// SIMATIC S7-200 project (STEP 7-Micro/WIN), CPU 224XP CN REL 02.01

ORGANIZATION_BLOCK MAIN:OB1
TITLE=REALIZADO POR: BISMARK CHOQUE CHOQUE - REALIMENTACION DE ESTADOS
BEGIN
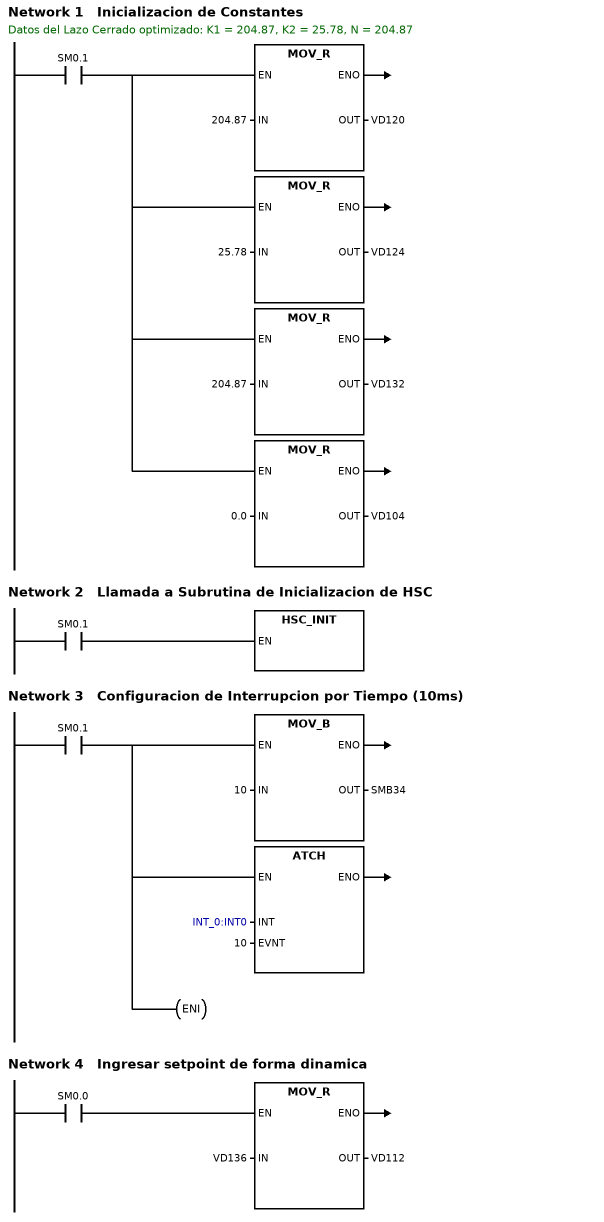
Network 1 //  Inicializacion de Constantes 
//  Datos del Lazo Cerrado optimizado: K1 = 204.87, K2 = 25.78, N = 204.87
// TU GANANCIA K1 (Posición)
// TU GANANCIA K2 (Velocidad)
// TU GANANCIA N (Pre-compensación calculada)
// Inicializar Pos_Anterior en 0.0
LD     SM0.1
MOVR   204.87, VD120
MOVR   25.78, VD124
MOVR   204.87, VD132
MOVR   0.0, VD104
Network 2 //  Llamada a Subrutina de Inicializacion de HSC
// Llamada a HSC_INIT
LD     SM0.1
CALL   HSC_INIT:SBR1
Network 3 //  Configuracion de Interrupcion por Tiempo (10ms)
// Intervalo de tiempo = 10 ms
// Asociar INT0 al evento de tiempo de SMB34
// Habilitar interrupciones globales
LD     SM0.1
MOVB   10, SMB34
ATCH   INT_0:INT0, 10
ENI
Network 4 //  Ingresar setpoint de forma dinamica
// Mover Setpoint desde VD136 a VD112
LD     SM0.0
MOVR   VD136, VD112
END_ORGANIZATION_BLOCK

SUBROUTINE_BLOCK HSC_INIT:SBR1
TITLE=
BEGIN
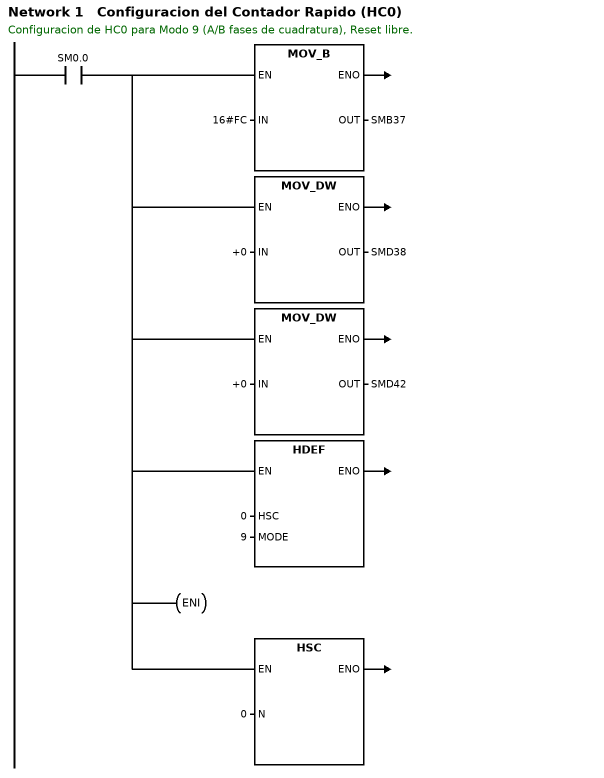
Network 1 //  Configuracion del Contador Rapido (HC0)
//  Configuracion de HC0 para Modo 9 (A/B fases de cuadratura), Reset libre.
// Control bits: Dirección arriba; escala 1X; habilitado
// Cargar valor actual en 0
// Cargar valor de preselección en 0
// Definir HC0 en Modo 9
// Asegurar habilitación de interrupciones
// Arrancar el contador rápido HC0
LD     SM0.0
MOVB   16#FC, SMB37
MOVD   +0, SMD38
MOVD   +0, SMD42
HDEF   0, 9
ENI
HSC    0
END_SUBROUTINE_BLOCK

INTERRUPT_BLOCK INT_0:INT0
TITLE=
BEGIN
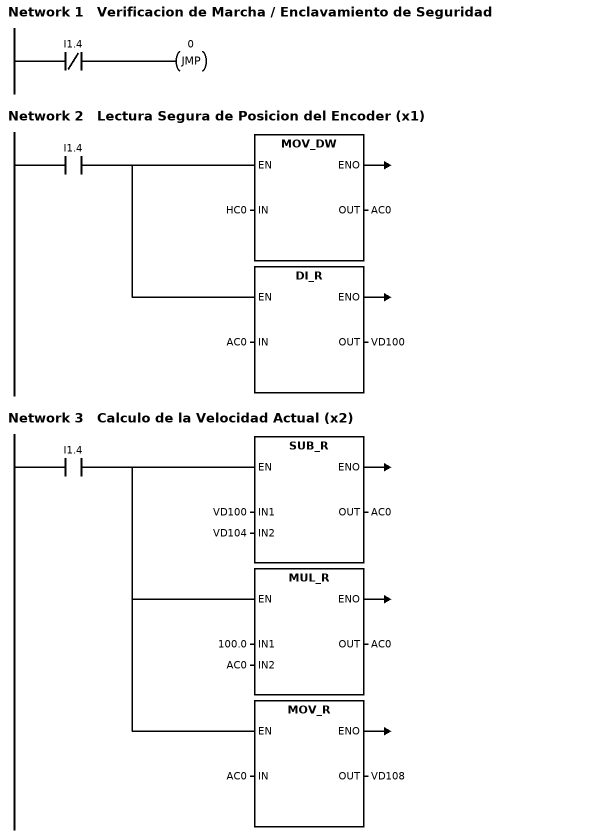
Network 1 //  Verificacion de Marcha / Enclavamiento de Seguridad
// Si I1.4 está desactivado (Emergencia/Stop)
// Salta directo a la parada segura (LBL 0)
LDN    I1.4
JMP    0
Network 2 //  Lectura Segura de Posicion del Encoder (x1)
// Leer cuentas acumuladas del hardware a AC0
// Convertir cuentas DINT a flotante REAL (x1)
LD     I1.4
MOVD   HC0, AC0
DTR    AC0, VD100
Network 3 //  Calculo de la Velocidad Actual (x2)
// Cuentas actuales
// Delta Posición = Cuentas_Actuales - Cuentas_Anteriores
// Delta_Pos / 0.01s equivale a multiplicar por 100.0
// Guardar en VD108 = Velocidad actual (x2)
LD     I1.4
MOVR   VD100, AC0
-R     VD104, AC0
*R     100.0, AC0
MOVR   AC0, VD108
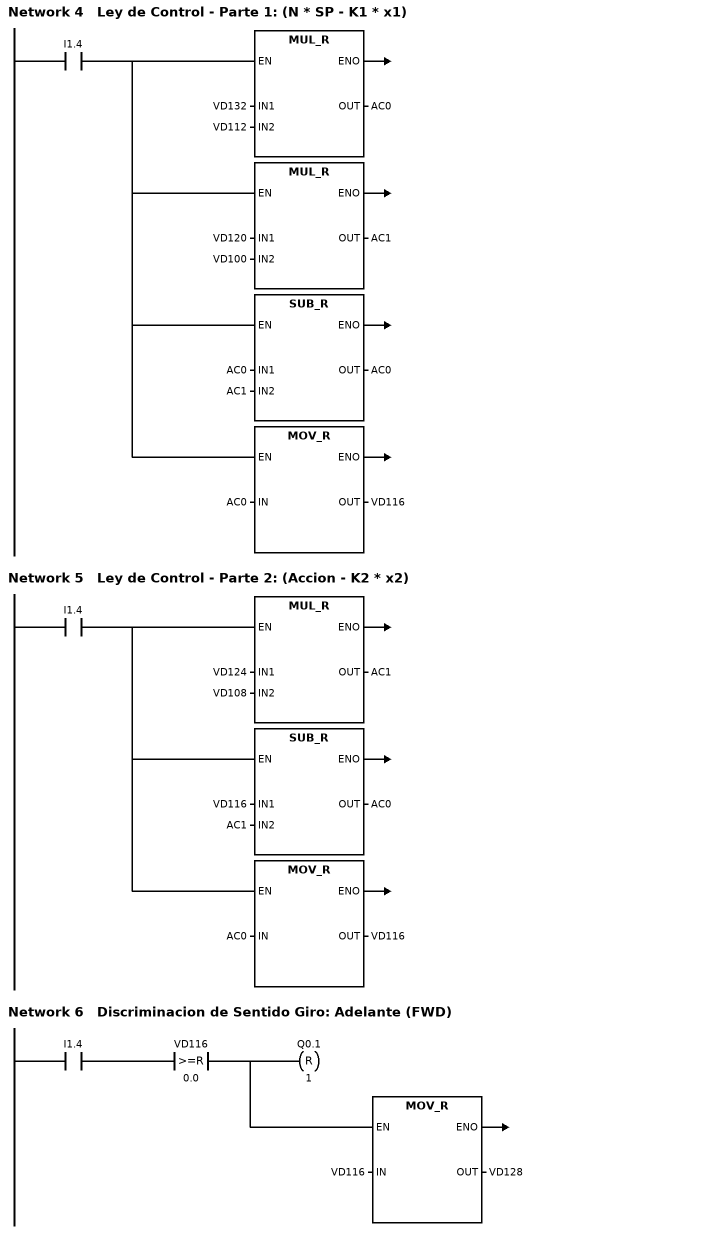
Network 4 //  Ley de Control - Parte 1: (N * SP - K1 * x1)
// Cargar N (204.87)
// AC0 = N * Setpoint
// Cargar K1 (204.87)
// AC1 = K1 * x1 (Posición)
// AC0 = (N * SP) - (K1 * x1)
// Almacenamiento intermedio
LD     I1.4
MOVR   VD132, AC0
*R     VD112, AC0
MOVR   VD120, AC1
*R     VD100, AC1
-R     AC1, AC0
MOVR   AC0, VD116
Network 5 //  Ley de Control - Parte 2: (Accion - K2 * x2)
// Cargar K2 (25.78)
// AC1 = K2 * x2 (Velocidad)
// Recuperar parte 1
// AC0 = (N * SP) - (K1 * x1) - (K2 * x2)
// VD116 = Acción de Control Final calculada (u)
LD     I1.4
MOVR   VD124, AC1
*R     VD108, AC1
MOVR   VD116, AC0
-R     AC1, AC0
MOVR   AC0, VD116
Network 6 //  Discriminacion de Sentido Giro: Adelante (FWD)
// Si u[k] es positiva o cero
// Desactivar salida de dirección reversa (Giro FWD)
// Guardar valor para magnitud |u|
LD     I1.4
AR>=   VD116, 0.0
R      Q0.1, 1
MOVR   VD116, VD128
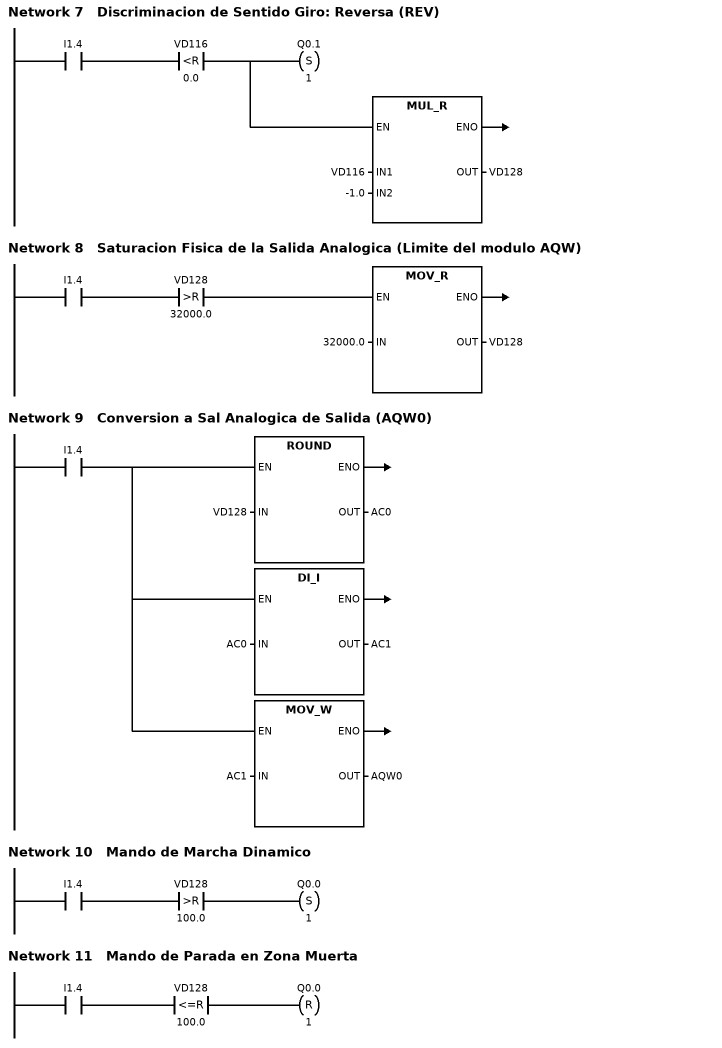
Network 7 //  Discriminacion de Sentido Giro: Reversa (REV)
// Si u[k] es negativa
// Activar salida física Q0.1 (Giro REV)
// Cargar u[k]
// Invertir signo para obtener valor absoluto |u|
LD     I1.4
AR<    VD116, 0.0
S      Q0.1, 1
MOVR   VD116, VD128
*R     -1.0, VD128
Network 8 //  Saturacion Fisica de la Salida Analogica (Limite del modulo AQW)
// Si excede el límite del módulo analógico de Siemens
// Recortar la acción a un máximo de 32000 unidades
LD     I1.4
AR>    VD128, 32000.0
MOVR   32000.0, VD128
Network 9 //  Conversion a Sal Analogica de Salida (AQW0)
// Convertir de flotante REAL a DINT
// Convertir de DINT a entero de 16 bits INT
// Enviar el valor numérico al canal físico del Variador
LD     I1.4
ROUND  VD128, AC0
DTI    AC0, AC1
MOVW   AC1, AQW0
Network 10 //  Mando de Marcha Dinamico
// Si hay suficiente tensión asignada (evita zumbidos)
// Energizar el contactor de marcha / habilitación
LD     I1.4
AR>    VD128, 100.0
S      Q0.0, 1
Network 11 //  Mando de Parada en Zona Muerta
// Si la acción es prácticamente cero
// Apagar la habilitación del motor
LD     I1.4
AR<=   VD128, 100.0
R      Q0.0, 1
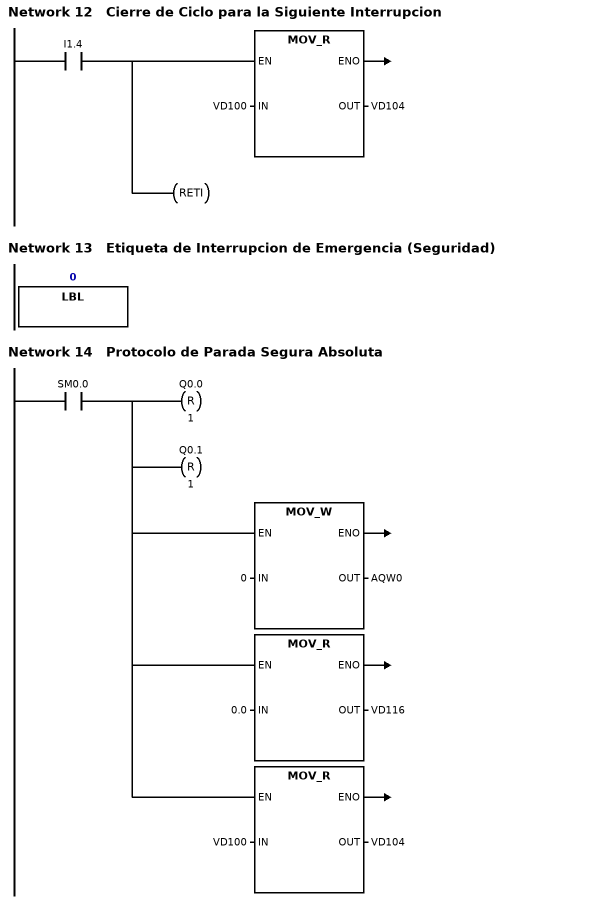
Network 12 //  Cierre de Ciclo para la Siguiente Interrupcion
// Pos_Anterior = Pos_Actual
// Retorno condicional de la interrupción
LD     I1.4
MOVR   VD100, VD104
CRETI
Network 13 //  Etiqueta de Interrupcion de Emergencia (Seguridad)
LBL    0
Network 14 //  Protocolo de Parada Segura Absoluta
// Desactivar salida de Marcha
// Desactivar salida de Dirección
// Forzar voltaje del variador a 0V
// Vaciar registro de control
// Sincronizar estados para evitar saltos bruscos al volver
LD     SM0.0
R      Q0.0, 1
R      Q0.1, 1
MOVW   0, AQW0
MOVR   0.0, VD116
MOVR   VD100, VD104
END_INTERRUPT_BLOCK
